Yaskawa INFORM job: BASIC-W-ARC-GAJ.JBI

/JOB
//NAME BASIC-W-ARC-GAJ
///FOLDERNAME GABEJ-YRC1000
//POS
///NPOS 14,0,14,1,0,1
///TOOL 0
///POSTYPE PULSE
///PULSE
C00000=4452,18827,-51072,2986,-34195,44008
C00001=765,27316,-49630,10024,-29036,41831
C00002=-3236,40072,-26608,5060,-37172,18423
C00003=-14145,43687,-19462,11285,-41287,-18176
C00004=-15498,47150,-14668,9494,-47224,-18653
C00005=-15777,47283,-12103,9236,-48386,-18239
C00006=-23740,8119,-77161,5340,15629,-8173
C00007=-20127,15447,-75197,-11658,16665,-481
C00008=-22177,16500,-71146,27954,10527,-20920
C00009=-19671,9683,-70517,8540,5629,-10803
C00010=-25009,7130,-105405,782,47608,-17190
C00011=-22296,10885,-88726,-1645,23061,-16261
C00012=-20888,15802,-83207,-3273,22976,-15885
C00013=-23771,9748,-100031,-181,45881,-17086
EC00000=-12851
EC00001=-1530
EC00002=-1510
EC00003=-2717
EC00004=-2717
EC00005=-3439
EC00006=-82435
EC00007=-82434
EC00008=-82435
EC00009=-82435
EC00010=-160520
EC00011=-150746
EC00012=-150746
EC00013=-160520
P00100=0,-60000,-60000,0,-90000,0
EX00100=0
//INST
///DATE 2026/08/06 16:48
///ATTR SC,RW
///GROUP1 RB1,ST1
NOP
MOVJ P100 EX100 VJ=5.00
MOVJ C00000 EC00000 VJ=50.00
MOVC C00001 EC00001 V=83.3
ARCON ASF#(14)
WVON WEV#(12)
MOVC C00002 EC00002
MOVC C00003 EC00003
MOVC C00004 EC00004 FPT
WVOF
ARCOF AEF#(12)
MOVL C00005 EC00005 V=83.3
MOVJ C00006 EC00006 VJ=25.00
MOVL C00007 EC00007 V=83.3
ARCON ASF#(12)
WVON WEV#(12)
MOVL C00008 EC00008
WVOF
ARCOF AEF#(12)
MOVL C00009 EC00009 V=333.3
MOVL C00010 EC00010 V=333.3
MOVL C00011 EC00011 V=50.0
ARCON ASF#(13)
COMM WVON WEV#(12)
MOVL C00012 EC00012
WVOF
ARCOF AEF#(13)
MOVL C00013 EC00013 V=333.3
MOVJ P100 EX100 VJ=50.00
CALL JOB:CLEAN_R1
END
